Staubli VAL3: changeDataLib1.pgx

public program changeDataLib1(num x_nLib (dimensions=1))
  local num l_nClock
  local num l_nResult
begin
  //形参：x_nLib
  //对应实参：savedata:nLibIndex
  //  bTosave=true
  //  call trajectory:onSave(bTosave)
  //  bTosave=true
  //  call prog:onSave(bTosave)
  l_nClock=clock()
  logMsg("自动开始切换库:"+toString(".2",clock()))
  call trajectory:loadTRAJ(x_nLib,l_nResult)
  call prog:loadPROG(x_nLib,l_nResult)

  delay(1)
  logMsg(toString(".3",clock()-l_nClock))
end
